Fanuc KAREL source: kd00058.KL

-- PROVISIONAL review KL for V1013-1; original PC SHA256 dab9e8e52811d95e46284d54452878e38f3c36d3a25b56ec42a8820feb82e867
-- Incomplete behavior may be omitted. Consult companion uncertainty JSON. Do not deploy.
PROGRAM KD00058
%NOLOCKGROUP
VAR
  I : INTEGER
  J : INTEGER
  B : BOOLEAN
  R : REAL
  S : STRING[80]
BEGIN
  -- UNRESOLVED_PC offsets 5-18; opcodes 9D,81,18,9D,1B,9D,12,9C,13,04
  -- UNRESOLVED_PC offsets 23-27; opcodes 7F
END KD00058
